(* IEC 61131-3 sources: PLCGen/codesys_service/bank/custom/st, 12 files *)

(* ---- FB_C01.st ---- *)
FUNCTION_BLOCK FB_C01
VAR_INPUT
    RunSwitch : BOOL;
    PartPresent : BOOL;
    DefectSensor : BOOL;
    ResetButton : BOOL;
END_VAR
VAR_OUTPUT
    ConveyorMotor : BOOL;
    RejectPusher : BOOL;
    AcceptCount : INT;
    RejectCount : INT;
    BatchFull : BOOL;
END_VAR
VAR
    prevPart : BOOL;
    partEdge : BOOL;
    rejectPulse : BOOL;
    pusherTimer : TOF;
    total : INT;
END_VAR

partEdge := PartPresent AND NOT prevPart;
rejectPulse := partEdge AND DefectSensor AND RunSwitch AND NOT BatchFull;
pusherTimer(IN := rejectPulse, PT := T#1S);

IF ResetButton THEN
    AcceptCount := 0;
    RejectCount := 0;
    BatchFull := FALSE;
ELSIF partEdge AND RunSwitch AND NOT BatchFull THEN
    IF DefectSensor THEN
        RejectCount := RejectCount + 1;
    ELSE
        AcceptCount := AcceptCount + 1;
    END_IF;
    total := AcceptCount + RejectCount;
    IF total >= 5 THEN
        BatchFull := TRUE;
    END_IF;
END_IF;

ConveyorMotor := RunSwitch AND NOT BatchFull;
RejectPusher := pusherTimer.Q AND NOT BatchFull;
prevPart := PartPresent;

(* ---- FB_C02.st ---- *)
FUNCTION_BLOCK FB_C02
VAR_INPUT
    LeftButton : BOOL;
    RightButton : BOOL;
    PartPresent : BOOL;
    ResetButton : BOOL;
END_VAR
VAR_OUTPUT
    PressOutput : BOOL;
    CycleComplete : BOOL;
    Fault : BOOL;
END_VAR
VAR
    leftTimer : TON;
    rightTimer : TON;
    pressWasOn : BOOL;
END_VAR

leftTimer(IN := LeftButton AND NOT RightButton, PT := T#500MS);
rightTimer(IN := RightButton AND NOT LeftButton, PT := T#500MS);

IF leftTimer.Q OR rightTimer.Q THEN
    Fault := TRUE;
END_IF;

IF ResetButton AND NOT LeftButton AND NOT RightButton THEN
    Fault := FALSE;
END_IF;

PressOutput := LeftButton AND RightButton AND PartPresent AND NOT Fault;
CycleComplete := pressWasOn AND NOT PressOutput;
pressWasOn := PressOutput;

(* ---- FB_C03.st ---- *)
FUNCTION_BLOCK FB_C03
VAR_INPUT
    VehiclePresent : BOOL;
    OpenButton : BOOL;
    SafetyBeam : BOOL;
END_VAR
VAR_OUTPUT
    GateOpen : BOOL;
    GateClosed : BOOL;
    WarningLight : BOOL;
END_VAR
VAR
    gateOpenState : BOOL;
    prevOpenButton : BOOL;
    closeTimer : TON;
END_VAR

IF ((OpenButton AND NOT prevOpenButton) OR VehiclePresent OR SafetyBeam) THEN
    gateOpenState := TRUE;
END_IF;

closeTimer(IN := gateOpenState AND NOT VehiclePresent AND NOT SafetyBeam AND NOT OpenButton, PT := T#3S);
IF closeTimer.Q THEN
    gateOpenState := FALSE;
END_IF;

GateOpen := gateOpenState;
GateClosed := NOT gateOpenState;
WarningLight := SafetyBeam;
prevOpenButton := OpenButton;

(* ---- FB_C04.st ---- *)
FUNCTION_BLOCK FB_C04
VAR_INPUT
    StartButton : BOOL;
    StopButton : BOOL;
    Overload : BOOL;
    ResetButton : BOOL;
END_VAR
VAR_OUTPUT
    MainContactor : BOOL;
    StarContactor : BOOL;
    DeltaContactor : BOOL;
    Running : BOOL;
    Fault : BOOL;
END_VAR
VAR
    prevStart : BOOL;
    startEdge : BOOL;
    starTimer : TON;
END_VAR

startEdge := StartButton AND NOT prevStart;

IF Overload THEN
    Fault := TRUE;
END_IF;
IF ResetButton AND NOT Overload THEN
    Fault := FALSE;
END_IF;

IF Fault OR StopButton THEN
    MainContactor := FALSE;
    StarContactor := FALSE;
    DeltaContactor := FALSE;
    Running := FALSE;
    starTimer(IN := FALSE, PT := T#3S);
ELSIF startEdge THEN
    MainContactor := TRUE;
    StarContactor := TRUE;
    DeltaContactor := FALSE;
    Running := TRUE;
    starTimer(IN := TRUE, PT := T#3S);
ELSE
    IF MainContactor THEN
        starTimer(IN := StarContactor, PT := T#3S);
        IF starTimer.Q THEN
            StarContactor := FALSE;
            DeltaContactor := TRUE;
        END_IF;
    END_IF;
END_IF;

prevStart := StartButton;

(* ---- FB_C05.st ---- *)
FUNCTION_BLOCK FB_C05
VAR_INPUT
    StartButton : BOOL;
    EmergencyStop : BOOL;
    VehiclePresent : BOOL;
    ResetButton : BOOL;
END_VAR
VAR_OUTPUT
    ConveyorMotor : BOOL;
    FoamValve : BOOL;
    BrushMotor : BOOL;
    RinseValve : BOOL;
    DryFan : BOOL;
    CycleComplete : BOOL;
    Fault : BOOL;
END_VAR
VAR
    step : INT;
    prevStart : BOOL;
    startEdge : BOOL;
    foamTimer : TON;
    brushTimer : TON;
    rinseTimer : TON;
    dryTimer : TON;
END_VAR

startEdge := StartButton AND NOT prevStart;
foamTimer(IN := (step = 1), PT := T#2S);
brushTimer(IN := (step = 2), PT := T#2S);
rinseTimer(IN := (step = 3), PT := T#1S);
dryTimer(IN := (step = 4), PT := T#1S);

IF EmergencyStop THEN
    Fault := TRUE;
    step := 0;
END_IF;
IF ResetButton THEN
    Fault := FALSE;
    CycleComplete := FALSE;
END_IF;

IF startEdge AND VehiclePresent AND NOT Fault AND NOT EmergencyStop THEN
    step := 1;
    CycleComplete := FALSE;
END_IF;

IF step = 1 AND foamTimer.Q THEN
    step := 2;
END_IF;
IF step = 2 AND brushTimer.Q THEN
    step := 3;
END_IF;
IF step = 3 AND rinseTimer.Q THEN
    step := 4;
END_IF;
IF step = 4 AND dryTimer.Q THEN
    step := 5;
END_IF;
IF step = 5 THEN
    step := 0;
    CycleComplete := TRUE;
END_IF;

ConveyorMotor := (step >= 1) AND (step <= 4) AND NOT EmergencyStop AND NOT Fault;
FoamValve := (step = 1) AND NOT EmergencyStop AND NOT Fault;
BrushMotor := (step = 2) AND NOT EmergencyStop AND NOT Fault;
RinseValve := (step = 3) AND NOT EmergencyStop AND NOT Fault;
DryFan := (step = 4) AND NOT EmergencyStop AND NOT Fault;
prevStart := StartButton;

(* ---- FB_C06.st ---- *)
FUNCTION_BLOCK FB_C06
VAR_INPUT
    OpenButton : BOOL;
    CloseButton : BOOL;
    ObstacleSensor : BOOL;
    DoorOpenLimit : BOOL;
    DoorClosedLimit : BOOL;
    ResetButton : BOOL;
END_VAR
VAR_OUTPUT
    DoorMotorOpen : BOOL;
    DoorMotorClose : BOOL;
    DoorOpen : BOOL;
    DoorClosed : BOOL;
    WarningBuzzer : BOOL;
    Fault : BOOL;
END_VAR
VAR
    opening : BOOL;
    closing : BOOL;
    autoTimer : TON;
END_VAR

IF DoorOpenLimit AND DoorClosedLimit THEN
    Fault := TRUE;
    opening := FALSE;
    closing := FALSE;
ELSIF ResetButton THEN
    Fault := FALSE;
END_IF;

IF NOT Fault THEN
    IF (OpenButton AND NOT DoorOpenLimit) OR (ObstacleSensor AND closing) THEN
        opening := TRUE;
        closing := FALSE;
    END_IF;

    IF CloseButton AND NOT ObstacleSensor AND NOT OpenButton THEN
        closing := TRUE;
        opening := FALSE;
    END_IF;

    autoTimer(IN := DoorOpenLimit AND NOT ObstacleSensor AND NOT OpenButton AND NOT CloseButton, PT := T#5S);
    IF autoTimer.Q AND NOT ObstacleSensor THEN
        closing := TRUE;
        opening := FALSE;
    END_IF;

    IF ObstacleSensor THEN
        opening := TRUE;
        closing := FALSE;
    END_IF;

    IF opening AND DoorOpenLimit THEN
        opening := FALSE;
    END_IF;
    IF closing AND DoorClosedLimit THEN
        closing := FALSE;
    END_IF;
ELSE
    opening := FALSE;
    closing := FALSE;
    autoTimer(IN := FALSE, PT := T#5S);
END_IF;

DoorMotorOpen := opening;
DoorMotorClose := closing;
DoorOpen := DoorOpenLimit;
DoorClosed := DoorClosedLimit;
WarningBuzzer := ObstacleSensor;

(* ---- FB_C07.st ---- *)
FUNCTION_BLOCK FB_C07
VAR_INPUT
    RunSwitch : BOOL;
    PartPresent : BOOL;
    HeightSensor : REAL;
    ResetButton : BOOL;
END_VAR
VAR_OUTPUT
    ConveyorMotor : BOOL;
    AcceptGate : BOOL;
    RejectGate : BOOL;
    AcceptCount : INT;
    RejectCount : INT;
    Fault : BOOL;
END_VAR
VAR
    prevPart : BOOL;
    partEdge : BOOL;
    acceptPulse : BOOL;
    rejectPulse : BOOL;
    acceptTimer : TOF;
    rejectTimer : TOF;
END_VAR

IF (HeightSensor < 0.0) OR (HeightSensor > 100.0) THEN
    Fault := TRUE;
END_IF;
IF ResetButton THEN
    AcceptCount := 0;
    RejectCount := 0;
    Fault := FALSE;
END_IF;

partEdge := PartPresent AND NOT prevPart;
acceptPulse := partEdge AND RunSwitch AND NOT Fault AND (HeightSensor >= 40.0) AND (HeightSensor <= 60.0);
rejectPulse := partEdge AND RunSwitch AND NOT Fault AND ((HeightSensor < 40.0) OR (HeightSensor > 60.0));

acceptTimer(IN := acceptPulse, PT := T#500MS);
rejectTimer(IN := rejectPulse, PT := T#500MS);
AcceptGate := acceptTimer.Q;
RejectGate := rejectTimer.Q;

IF acceptPulse THEN
    AcceptCount := AcceptCount + 1;
ELSIF rejectPulse THEN
    RejectCount := RejectCount + 1;
END_IF;

ConveyorMotor := RunSwitch AND NOT Fault;
prevPart := PartPresent;

(* ---- FB_C08.st ---- *)
FUNCTION_BLOCK FB_C08
VAR_INPUT
    StartButton : BOOL;
    StopButton : BOOL;
    Zone1Moisture : REAL;
    Zone2Moisture : REAL;
    Zone3Moisture : REAL;
    ResetButton : BOOL;
END_VAR
VAR_OUTPUT
    Zone1Valve : BOOL;
    Zone2Valve : BOOL;
    Zone3Valve : BOOL;
    Pump : BOOL;
    CycleComplete : BOOL;
END_VAR
VAR
    step : INT;
    prevStart : BOOL;
    startEdge : BOOL;
    zone1Timer : TON;
    zone2Timer : TON;
    zone3Timer : TON;
END_VAR

startEdge := StartButton AND NOT prevStart;
zone1Timer(IN := (step = 1) AND (Zone1Moisture < 30.0), PT := T#3S);
zone2Timer(IN := (step = 2) AND (Zone2Moisture < 30.0), PT := T#3S);
zone3Timer(IN := (step = 3) AND (Zone3Moisture < 30.0), PT := T#3S);

IF StopButton THEN
    step := 0;
    CycleComplete := FALSE;
END_IF;
IF ResetButton THEN
    CycleComplete := FALSE;
END_IF;
IF startEdge AND NOT CycleComplete AND NOT StopButton THEN
    step := 1;
    CycleComplete := FALSE;
END_IF;

IF step = 1 AND Zone1Moisture >= 30.0 THEN
    step := 2;
END_IF;
IF step = 2 AND Zone2Moisture >= 30.0 THEN
    step := 3;
END_IF;
IF step = 3 AND Zone3Moisture >= 30.0 THEN
    step := 4;
END_IF;
IF (zone1Timer.Q OR zone2Timer.Q OR zone3Timer.Q) THEN
    step := step + 1;
END_IF;
IF step = 4 THEN
    step := 0;
    CycleComplete := TRUE;
END_IF;

Zone1Valve := (step = 1) AND (Zone1Moisture < 30.0) AND NOT StopButton;
Zone2Valve := (step = 2) AND (Zone2Moisture < 30.0) AND NOT StopButton;
Zone3Valve := (step = 3) AND (Zone3Moisture < 30.0) AND NOT StopButton;
Pump := Zone1Valve OR Zone2Valve OR Zone3Valve;
prevStart := StartButton;

(* ---- FB_C09.st ---- *)
FUNCTION_BLOCK FB_C09
VAR_INPUT
    RunSwitch : BOOL;
    Zone1Sensor : BOOL;
    Zone2Sensor : BOOL;
    Zone3Sensor : BOOL;
    ReleaseButton : BOOL;
    ResetButton : BOOL;
END_VAR
VAR_OUTPUT
    Zone1Motor : BOOL;
    Zone2Motor : BOOL;
    Zone3Motor : BOOL;
    Zone1Full : BOOL;
    Zone2Full : BOOL;
    Zone3Full : BOOL;
    JamAlarm : BOOL;
END_VAR
VAR
    z1Timer : TON;
    z2Timer : TON;
    z3Timer : TON;
END_VAR

IF ResetButton THEN
    JamAlarm := FALSE;
END_IF;

Zone3Motor := RunSwitch AND Zone3Sensor AND ReleaseButton;
Zone2Motor := RunSwitch AND Zone2Sensor AND NOT Zone3Sensor;
Zone1Motor := RunSwitch AND Zone1Sensor AND NOT Zone2Sensor;

Zone1Full := Zone1Sensor AND Zone2Sensor;
Zone2Full := Zone2Sensor AND Zone3Sensor;
Zone3Full := Zone3Sensor AND NOT ReleaseButton;

z1Timer(IN := RunSwitch AND Zone1Sensor AND NOT Zone1Motor, PT := T#5S);
z2Timer(IN := RunSwitch AND Zone2Sensor AND NOT Zone2Motor, PT := T#5S);
z3Timer(IN := RunSwitch AND Zone3Sensor AND NOT Zone3Motor, PT := T#5S);

IF z1Timer.Q OR z2Timer.Q OR z3Timer.Q THEN
    JamAlarm := TRUE;
END_IF;

IF JamAlarm THEN
    Zone1Motor := FALSE;
    Zone2Motor := FALSE;
    Zone3Motor := FALSE;
END_IF;

(* ---- FB_C10.st ---- *)
FUNCTION_BLOCK FB_C10
VAR_INPUT
    StartButton : BOOL;
    StopButton : BOOL;
    EmergencyStop : BOOL;
    FlameSensor : BOOL;
    ResetButton : BOOL;
END_VAR
VAR_OUTPUT
    PurgeFan : BOOL;
    Igniter : BOOL;
    FuelValve : BOOL;
    FlameOn : BOOL;
    Lockout : BOOL;
    Fault : BOOL;
END_VAR
VAR
    step : INT;
    prevStart : BOOL;
    startEdge : BOOL;
    purgeTimer : TON;
    igniteTimer : TON;
END_VAR

startEdge := StartButton AND NOT prevStart;
purgeTimer(IN := (step = 1), PT := T#3S);
igniteTimer(IN := (step = 2), PT := T#2S);

IF EmergencyStop THEN
    Fault := TRUE;
    step := 0;
END_IF;
IF StopButton THEN
    step := 0;
END_IF;
IF ResetButton AND NOT StartButton AND NOT FlameSensor THEN
    Lockout := FALSE;
    Fault := FALSE;
END_IF;
IF startEdge AND NOT Lockout AND NOT Fault AND NOT EmergencyStop THEN
    step := 1;
END_IF;

IF step = 1 AND purgeTimer.Q THEN
    step := 2;
END_IF;
IF step = 2 THEN
    IF FlameSensor THEN
        step := 3;
    ELSIF igniteTimer.Q THEN
        Lockout := TRUE;
        step := 0;
    END_IF;
END_IF;
IF step = 3 AND NOT FlameSensor THEN
    Lockout := TRUE;
    step := 0;
END_IF;

FlameOn := (step = 3) AND FlameSensor;
PurgeFan := (step = 1) AND NOT EmergencyStop AND NOT Fault;
Igniter := (step = 2) AND NOT EmergencyStop AND NOT Fault;
FuelValve := (step = 3) AND FlameOn AND NOT EmergencyStop AND NOT StopButton AND NOT Fault;
prevStart := StartButton;

(* ---- FB_C11.st ---- *)
FUNCTION_BLOCK FB_C11
VAR_INPUT
    RunSwitch : BOOL;
    BoxPresent : BOOL;
    ResetButton : BOOL;
END_VAR
VAR_OUTPUT
    ConveyorMotor : BOOL;
    LayerPush : BOOL;
    BoxCount : INT;
    LayerCount : INT;
    PalletFull : BOOL;
END_VAR
VAR
    prevBox : BOOL;
    partEdge : BOOL;
    layerTrigger : BOOL;
    layerTimer : TOF;
END_VAR

partEdge := BoxPresent AND NOT prevBox;
layerTrigger := FALSE;

IF ResetButton THEN
    BoxCount := 0;
    LayerCount := 0;
    PalletFull := FALSE;
END_IF;

IF partEdge AND RunSwitch AND NOT PalletFull THEN
    BoxCount := BoxCount + 1;
END_IF;
IF BoxCount >= 3 THEN
    BoxCount := 0;
    LayerCount := LayerCount + 1;
    layerTrigger := TRUE;
END_IF;

layerTimer(IN := layerTrigger, PT := T#1S);
LayerPush := layerTimer.Q;

IF LayerCount >= 2 THEN
    PalletFull := TRUE;
END_IF;

ConveyorMotor := RunSwitch AND NOT PalletFull AND NOT LayerPush;
prevBox := BoxPresent;

(* ---- FB_C12.st ---- *)
FUNCTION_BLOCK FB_C12
VAR_INPUT
    RunSwitch : BOOL;
    LightCurtain : BOOL;
    MutingSensor1 : BOOL;
    MutingSensor2 : BOOL;
    ResetButton : BOOL;
END_VAR
VAR_OUTPUT
    ConveyorMotor : BOOL;
    MutingActive : BOOL;
    SafetyStop : BOOL;
    Alarm : BOOL;
END_VAR
VAR
    prevM1 : BOOL;
    prevM2 : BOOL;
    mutingArmed : BOOL;
    mutingActiveState : BOOL;
    muteWindow : TON;
END_VAR

muteWindow(IN := mutingArmed, PT := T#2S);

IF ResetButton AND NOT LightCurtain THEN
    SafetyStop := FALSE;
    Alarm := FALSE;
END_IF;

IF MutingSensor1 AND NOT prevM1 THEN
    mutingArmed := TRUE;
END_IF;

IF MutingSensor2 AND NOT prevM2 THEN
    IF mutingArmed AND NOT muteWindow.Q THEN
        mutingActiveState := TRUE;
    ELSE
        Alarm := TRUE;
    END_IF;
    mutingArmed := FALSE;
END_IF;

IF muteWindow.Q THEN
    Alarm := TRUE;
    mutingArmed := FALSE;
END_IF;

IF NOT (MutingSensor1 AND MutingSensor2) THEN
    mutingActiveState := FALSE;
END_IF;

IF LightCurtain AND NOT mutingActiveState THEN
    SafetyStop := TRUE;
END_IF;

ConveyorMotor := RunSwitch AND NOT SafetyStop AND (NOT LightCurtain OR mutingActiveState) AND NOT Alarm;
MutingActive := mutingActiveState;
prevM1 := MutingSensor1;
prevM2 := MutingSensor2;
